# EPICS autosave request: 1.5.0/debian-12/7.0.10/modules/ADCore-ee039d2/db/NDFileNexus_settings.req
$(P)$(R)TemplateFilePath
$(P)$(R)TemplateFileName
file "NDPluginFile_settings.req", P=$(P), R=$(R)
